Fanuc KAREL source: kt00473.KL

-- PROVISIONAL review KL for V1013-1; original PC SHA256 a2b367f2a35bd9a0ee7793f53347a9101d650c86cc6e94d72b60ee94d2017e56
-- Incomplete behavior may be omitted. Consult companion uncertainty JSON. Do not deploy.
PROGRAM KT00473
%NOLOCKGROUP
VAR
  OUT : BOOLEAN
-- UNRESOLVED_DECL P1 type=000101
-- UNRESOLVED_DECL P2 type=000101
BEGIN
  -- UNRESOLVED_PC offsets 5-28; opcodes 49,49,AC,23
  -- UNRESOLVED_PC offsets 33-37; opcodes 7F
END KT00473
